// TIA Portal V20 export
// export: Created 2026-10-20T12:46:10.4769616Z, ExportSetting WithDefaults, DisplayName Totally Integrated Automation Portal, DisplayVersion V20 Update 6, DisplayName TIA Portal Openness, DisplayVersion V20 Update 6, DisplayName TIA Portal Version Control Interface, DisplayVersion V20 Update 6, DisplayName SINAMICS Startdrive Advanced, DisplayVersion V20 SP1, DisplayName SINAMICS Startdrive G130, G150, S120, S150, SINAMICS MV, G220, S200, S210, DisplayVersion V20 SP1, DisplayName SINAMICS Startdrive G110M, G120, G120C, G120D, G120P, G115D, DisplayVersion V20 SP1, DisplayName STEP 7 Professional, DisplayVersion V20 Update 6, DisplayName STEP 7 Safety, DisplayVersion V20 Update 2, DisplayName WinCC Basic/Comfort/Advanced, DisplayVersion V20 Update 6, DisplayName WinCC Unified, DisplayVersion V20 Update 6
DATA_BLOCK "Screen_DB"   // DB23
{ S7_Optimized_Access := 'TRUE' }
VERSION : 0.1
// stored: AutoNumber true, DBAccessibleFromOPCUA true, IsOnlyStoredInLoadMemory false, IsRetainMemResEnabled false, IsWriteProtectedInAS false, MemoryReserve 100
   VAR
      Settings_ActivePopUp : USInt;
      Alarms_ActiveTable : USInt;
      MainTemplate_ErrorActive : Bool;
      MainTemplate_ErrorCount : USInt;
      MainTemplate_Background : USInt;
      EmptyTemplate_Background : USInt;
      Charge_VTD : Bool;
      Charge_Cnv : Bool;
      Charge_VTD_Commands : Bool;
      Charge_Cnv_Commands : Bool;
      Charge_OT : Bool;
      Shuttle : "Shuttle_MQTT_Status_Msg";
      Shuttle_Select : USInt;
      VTD_Barcode : String;
      VTD_Barcode_Visu : Bool;
      OrderProcessing : Array[1..5] of String;
   END_VAR
BEGIN
END_DATA_BLOCK
